// TIA Portal V21 export
// export: Created 2026-11-21T13:24:04.6702441Z, ExportSetting WithDefaults, DisplayName Totally Integrated Automation Portal, DisplayVersion V21, DisplayName STEP 7 Professional, DisplayVersion V21, DisplayName STEP 7 Safety, DisplayVersion V21, DisplayName Tech WebApplication, DisplayVersion V21, DisplayName WinCC Basic/Comfort/Advanced, DisplayVersion V21, DisplayName WinCC Unified, DisplayVersion V21
FUNCTION_BLOCK "LineSafety"   // FB1, F_FBD
{ S7_Optimized_Access := 'TRUE' }
VERSION : 0.1
// Main safety block of the line's F-runtime group.
// stored: AutoNumber true, IsIECCheckEnabled false, UDAEnableTagReadback false
   VAR
      latched : Bool;
   END_VAR
BEGIN

REGION Network 1: Release
   // Released while start is pressed and the door is closed.
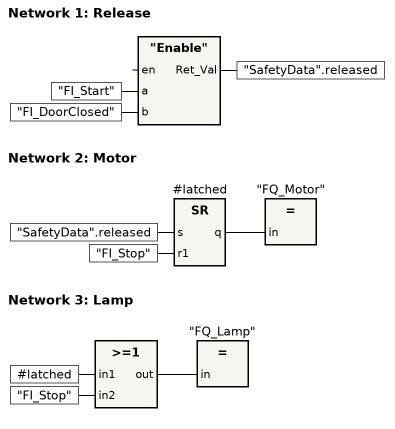
   "SafetyData".released := "Enable"("a" := "FI_Start", "b" := "FI_DoorClosed");
END_REGION

REGION Network 2: Motor
   // Latched on release, dropped by stop.
   IF "SafetyData".released THEN
       #latched := TRUE;   // SR flip-flop
   END_IF;
   IF "FI_Stop" THEN #latched := FALSE; END_IF;
   "FQ_Motor" := #latched;
END_REGION

REGION Network 3: Lamp
   // Lit while the motor runs or stop is pressed.
   "FQ_Lamp" := #latched OR "FI_Stop";
END_REGION
END_FUNCTION_BLOCK
